Fanuc KAREL source: kt00369.KL

-- PROVISIONAL review KL for V770-1; original PC SHA256 2e81aec0aa8df563ba2333357bdd7eaf52674d4ddd652e40ab0ad451494d5389
-- Incomplete behavior may be omitted. Consult companion uncertainty JSON. Do not deploy.
PROGRAM KT00369
%NOLOCKGROUP
VAR
  R1 : REAL
  I2 : INTEGER
  OUT : BOOLEAN
BEGIN
  -- UNRESOLVED_PC offsets 5-16; opcodes 2E,23
  -- UNRESOLVED_PC offsets 21-32; opcodes 2E,23
  -- UNRESOLVED_PC offsets 37-57; opcodes 21,21,64,70,23
  -- UNRESOLVED_PC offsets 62-66; opcodes 7F
END KT00369
